// TIA Portal V20 export
// export: Created 2026-10-19T18:07:28.5199214Z, ExportSetting WithDefaults, DisplayName Totally Integrated Automation Portal, DisplayVersion V20 Update 6, DisplayName TIA Portal Openness, DisplayVersion V20 Update 6, DisplayName TIA Portal Version Control Interface, DisplayVersion V20 Update 6, DisplayName SINAMICS Startdrive Advanced, DisplayVersion V20 SP1, DisplayName SINAMICS Startdrive G130, G150, S120, S150, SINAMICS MV, G220, S200, S210, DisplayVersion V20 SP1, DisplayName SINAMICS Startdrive G110M, G120, G120C, G120D, G120P, G115D, DisplayVersion V20 SP1, DisplayName STEP 7 Professional, DisplayVersion V20 Update 6, DisplayName STEP 7 Safety, DisplayVersion V20 Update 2, DisplayName WinCC Basic/Comfort/Advanced, DisplayVersion V20 Update 6, DisplayName WinCC Unified, DisplayVersion V20 Update 6
FUNCTION "ByteArrayToString_1" : String   // FC23, SCL
{ S7_Optimized_Access := 'TRUE' }
VERSION : 0.1
// stored: AutoNumber true, IsIECCheckEnabled false, SetENOAutomatically false, UDAEnableTagReadback false
   VAR_INPUT
      Lenght : Int;
      ByteArray : Array[1..200] of Byte;
   END_VAR
   VAR_TEMP
      tempStr_1 : String;
      foundPos : Int;
      i : Int;
   END_VAR
BEGIN
   #tempStr_1 := '';
   FOR #i := 1 TO MIN(IN1 := #Lenght - 1, IN2 := 200) DO
       IF #ByteArray[#i] <> 0 THEN
           #tempStr_1 := CONCAT(IN1 := #tempStr_1, IN2 := CHAR_TO_STRING(BYTE_TO_CHAR(#ByteArray[#i])));
       END_IF;
   END_FOR;

   // Remove '$02'
   // string 1
   #foundPos := FIND(IN1 := #tempStr_1, IN2 := '$02');
   WHILE #foundPos > 0 DO
       #tempStr_1 := REPLACE(IN1 := #tempStr_1, IN2 := '', P := #foundPos, L := 1);
       #foundPos := FIND(IN1 := #tempStr_1, IN2 := '$02');
   END_WHILE;

   #ByteArrayToString_1 := #tempStr_1;
END_FUNCTION
